(* IEC 61131-3 sources: OpenUnit/plc/lib/functions, 5 files *)

(* ---- FGEN5.st ---- *)
(* Function generator: piecewise linear f(X) through up to five points (X1,Y1)..(X5,Y5) with
   ascending X; constant beyond the end points.  For fewer points repeat the last one. *)
FUNCTION FGEN5 : REAL
  VAR_INPUT
    X : REAL;
    X1 : REAL;
    Y1 : REAL;
    X2 : REAL;
    Y2 : REAL;
    X3 : REAL;
    Y3 : REAL;
    X4 : REAL;
    Y4 : REAL;
    X5 : REAL;
    Y5 : REAL;
  END_VAR
  IF X <= X1 THEN
    FGEN5 := Y1;
  ELSIF X <= X2 THEN
    FGEN5 := Y1 + (Y2 - Y1) * (X - X1) / (X2 - X1);
  ELSIF X <= X3 THEN
    FGEN5 := Y2 + (Y3 - Y2) * (X - X2) / (X3 - X2);
  ELSIF X <= X4 THEN
    FGEN5 := Y3 + (Y4 - Y3) * (X - X3) / (X4 - X3);
  ELSIF X <= X5 THEN
    FGEN5 := Y4 + (Y5 - Y4) * (X - X4) / (X5 - X4);
  ELSE
    FGEN5 := Y5;
  END_IF;
END_FUNCTION

(* ---- FIRST_OUT.st ---- *)
(* First-out: number of the first TRUE input (C1 first), 0 when none is TRUE. The cause a first-out
   annunciator shows when several trip conditions come up in the same scan. Inputs left
   unconnected are FALSE. *)
FUNCTION FIRST_OUT : DINT
  VAR_INPUT
    C1 : BOOL := FALSE;
    C2 : BOOL := FALSE;
    C3 : BOOL := FALSE;
    C4 : BOOL := FALSE;
    C5 : BOOL := FALSE;
    C6 : BOOL := FALSE;
    C7 : BOOL := FALSE;
    C8 : BOOL := FALSE;
    C9 : BOOL := FALSE;
    C10 : BOOL := FALSE;
    C11 : BOOL := FALSE;
    C12 : BOOL := FALSE;
    C13 : BOOL := FALSE;
    C14 : BOOL := FALSE;
    C15 : BOOL := FALSE;
    C16 : BOOL := FALSE;
    C17 : BOOL := FALSE;
    C18 : BOOL := FALSE;
  END_VAR
  FIRST_OUT := 0;
  IF C18 THEN FIRST_OUT := 18; END_IF;
  IF C17 THEN FIRST_OUT := 17; END_IF;
  IF C16 THEN FIRST_OUT := 16; END_IF;
  IF C15 THEN FIRST_OUT := 15; END_IF;
  IF C14 THEN FIRST_OUT := 14; END_IF;
  IF C13 THEN FIRST_OUT := 13; END_IF;
  IF C12 THEN FIRST_OUT := 12; END_IF;
  IF C11 THEN FIRST_OUT := 11; END_IF;
  IF C10 THEN FIRST_OUT := 10; END_IF;
  IF C9 THEN FIRST_OUT := 9; END_IF;
  IF C8 THEN FIRST_OUT := 8; END_IF;
  IF C7 THEN FIRST_OUT := 7; END_IF;
  IF C6 THEN FIRST_OUT := 6; END_IF;
  IF C5 THEN FIRST_OUT := 5; END_IF;
  IF C4 THEN FIRST_OUT := 4; END_IF;
  IF C3 THEN FIRST_OUT := 3; END_IF;
  IF C2 THEN FIRST_OUT := 2; END_IF;
  IF C1 THEN FIRST_OUT := 1; END_IF;
END_FUNCTION

(* ---- MEDIAN3.st ---- *)
(* Median of three redundant transmitters (mid-value selection). *)
FUNCTION MEDIAN3 : REAL
  VAR_INPUT
    A : REAL;
    B : REAL;
    C : REAL;
  END_VAR
  MEDIAN3 := MAX(MIN(A, B), MIN(MAX(A, B), C));
END_FUNCTION

(* ---- TSAT.st ---- *)
(* Saturation temperature [degC] at pressure P [MPa abs] - IAPWS-IF97 derived table
   interpolated on ln(P), identical to tsat() in src/common/steamTable.js (generated from it). *)
FUNCTION TSAT : REAL
  VAR_INPUT
    P : REAL;
  END_VAR
  VAR
    PTAB : ARRAY[0..41] OF REAL := [0.001, 0.002, 0.003, 0.004, 0.005, 0.006, 0.008, 0.01, 0.015, 0.02, 0.03, 0.05, 0.07, 0.101325, 0.15, 0.2, 0.3, 0.5, 0.7, 1.0, 1.5, 2.0, 3.0, 4.0, 5.0, 6.0, 7.0, 8.0, 9.0, 10.0, 11.0, 12.0, 13.0, 14.0, 15.0, 16.0, 17.0, 18.0, 19.0, 20.0, 21.0, 21.8];
    TTAB : ARRAY[0..41] OF REAL := [6.97, 17.5, 24.08, 28.96, 32.88, 36.16, 41.51, 45.81, 53.97, 60.06, 69.1, 81.32, 89.95, 99.97, 111.35, 120.21, 133.52, 151.83, 164.95, 179.88, 198.29, 212.38, 233.86, 250.36, 263.94, 275.59, 285.83, 295.01, 303.35, 311.0, 318.08, 324.68, 330.86, 336.67, 342.16, 347.36, 352.29, 356.99, 361.47, 365.75, 369.83, 373.0];
    pc : REAL;
    x : REAL;
    i : INT;
    f : REAL;
  END_VAR
  pc := LIMIT(PTAB[0], P, PTAB[41]);
  x := LN(pc);
  i := 1;
  WHILE i < 41 AND LN(PTAB[i]) < x DO
    i := i + 1;
  END_WHILE;
  f := (x - LN(PTAB[i - 1])) / (LN(PTAB[i]) - LN(PTAB[i - 1]));
  TSAT := TTAB[i - 1] + f * (TTAB[i] - TTAB[i - 1]);
END_FUNCTION

(* ---- VOTE2OO3.st ---- *)
(* 2-out-of-3 voting of boolean trip channels. *)
FUNCTION VOTE2OO3 : BOOL
  VAR_INPUT
    A : BOOL;
    B : BOOL;
    C : BOOL;
  END_VAR
  VOTE2OO3 := (A AND B) OR (A AND C) OR (B AND C);
END_FUNCTION
